// Mitsubishi GX Works2 project: ABBACC   PLC: Q02/Q02H

PROGRAM MAIN
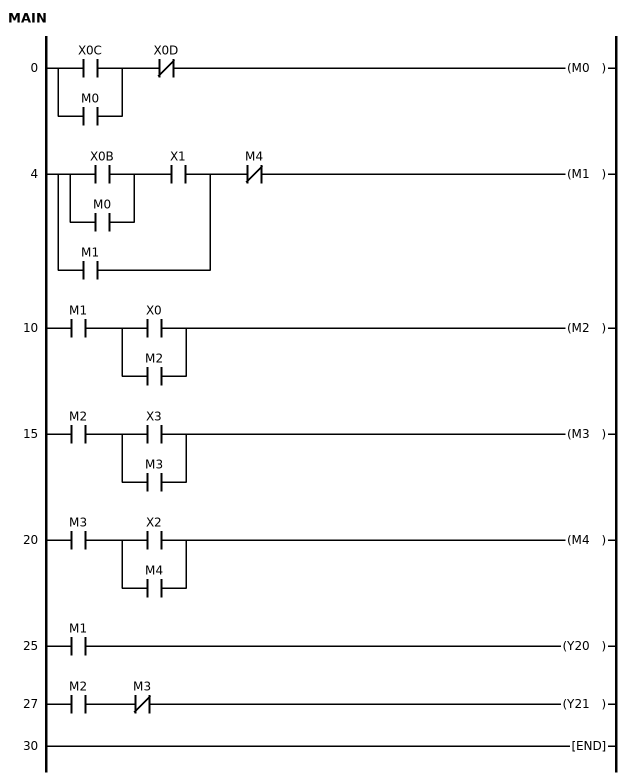
0     LD      X0C
      OR      M0
      ANI     X0D
      OUT     M0
4     LD      X0B
      OR      M0
      AND     X1
      OR      M1
      ANI     M4
      OUT     M1
10    LD      M1
      LD      X0
      OR      M2
      ANB
      OUT     M2
15    LD      M2
      LD      X3
      OR      M3
      ANB
      OUT     M3
20    LD      M3
      LD      X2
      OR      M4
      ANB
      OUT     M4
25    LD      M1
      OUT     Y20
27    LD      M2
      ANI     M3
      OUT     Y21
30    END
END_PROGRAM
